Staubli VAL3: updateTeachPos.pgx

public program updateTeachPos(point x_pteach, bool x_bteach)
begin
  if x_bteach==true
    utLbl_Point.Appearance.sBackgroundColour="#7CFA3F"
  else
    utLbl_Point.Appearance.sBackgroundColour="#FFFFFF"
  endIf
  utLbl_PosValue_Data[0].Common.sText=toString(".3",x_pteach.trsf.x)
  utLbl_PosValue_Data[1].Common.sText=toString(".3",x_pteach.trsf.y)
  utLbl_PosValue_Data[2].Common.sText=toString(".3",x_pteach.trsf.z)
  utLbl_PosValue_Data[3].Common.sText=toString(".3",x_pteach.trsf.rx)
  utLbl_PosValue_Data[4].Common.sText=toString(".3",x_pteach.trsf.ry)
  utLbl_PosValue_Data[5].Common.sText=toString(".3",x_pteach.trsf.rz)
end
